(* IEC 61131-3 sources: volt/packages/volt-lsp-iec/test-corpus/bakon-nano/Device/Plc Logic/Application/POUs/LenzeFunctions, 3 files *)

(* ---- SetRef_Axis.pou ---- *)
FUNCTION_BLOCK SetRef_Axis
VAR_INPUT
	I_AxisStatus	: KC_AxisBasicsStatus;
	I_lrHomeTarget	: LREAL;
END_VAR
VAR_OUTPUT
	Q_bRefDone		: BOOL;
	Q_bError		: BOOL;
END_VAR
VAR_IN_OUT
	IQ_CmdSetRef	: BOOL;
	IQ_Axis			: AXIS_REF;
	IQ_uControl_Axis	: KC_AxisBasicsControl;
END_VAR
VAR
	byStepper: BYTE;
	//LenzeECSWriteParameter1: L_DCO_ReadDriveParameter;
	bDone: BOOL;
	bError: BOOL;
	tWait: TON;
	//TestMultiturn: L_SMC_Multiturn;
	SetHomePosition : MC_SetPosition;
END_VAR

%LANGUAGE ST

CASE byStepper OF (*VERVALLEN, KAN NU VIA HOMING IN AXISBASICS: SET HOME -> SM3_Multiturn eronder aanroepen*)

	0:	Q_bRefDone							:=FALSE;
		Q_bError							:=FALSE;

		IF IQ_CmdSetRef
		THEN
			tWait(IN:= FALSE);
			IQ_uControl_Axis.bEnableDrive		:=FALSE;
			bDone								:=FALSE;
			bError								:=FALSE;
			IF NOT I_AxisStatus.bDriveEnabled THEN
				byStepper:=2;
			END_IF
		END_IF

	2:	SetHomePosition.Execute := TRUE;
		IF SetHomePosition.Done OR SetHomePosition.Error THEN
			byStepper := 4;
		END_IF

	4: Q_bRefDone := SetHomePosition.Done;
		Q_bError := SetHomePosition.Error;
		IF NOT IQ_CmdSetRef THEN
			byStepper := 0;
			SetHomePosition.Execute := FALSE;
		END_IF
END_CASE

SetHomePosition(
			Axis	:= IQ_Axis,
			Execute := ,
			Position:= I_lrHomeTarget,
			Relative	:= FALSE,
			Done=> ,
			Busy=> ,
			Error=> ,
			ErrorID=> );

END_FUNCTION_BLOCK

(* ---- XYA_MoveLineair_Bakon.pou ---- *)
(***********************************************************************************
Creation: LENL 		Datum: march 2008		Version: 1.0.0
 ***********************************************************************************
 FUNCTION:

FB for moving XYA in gear mode with a dummy axis. The dummy axis can be positioned or control external

 ***********************************************************************************
Name							Datum				Changes
Kling 							24.03.2009		Implementation

************************************************************************************
NOTE:

***********************************************************************************)

FUNCTION_BLOCK  XYA_MoveLineair_Bakon

VAR
	byStepper: BYTE;
	rMoveX: REAL;
	rMoveY: REAL;
	rMoveA: REAL;
	MC_GearIn_X: MC_GearIn;
	MC_GearIn_Y: MC_GearIn;
	MC_GearIn_A: MC_GearIn;
	MC_GearOut_X: MC_GearOut;
	MC_GearOut_Y: MC_GearOut;
	MC_GearOut_A: MC_GearOut;
	MC_MoveAbsolute_X: MC_MoveAbsolute;
	MC_MoveAbsolute_Y: MC_MoveAbsolute;
	MC_MoveAbsolute_A: MC_MoveAbsolute;
	CalcGearingRatio_X: CalcGearingRatio;
	CalcGearingRatio_Y: CalcGearingRatio;
	CalcGearingRatio_A: CalcGearingRatio;
	CalcGearingRatio_F: CalcGearingRatio;
	CalcGearingRatio_R: CalcGearingRatio;
	MC_MoveAbsolute_Mst: MC_MoveAbsolute;
	MC_SetPosition_Mst: MC_SetPosition;
	CalcMasterSpeedAcc_X: CalcMasterSpeedAcc;
	CalcMasterSpeedAcc_Y: CalcMasterSpeedAcc;
	CalcMasterSpeedAcc_A: CalcMasterSpeedAcc;
	CalcMasterSpeedAcc_F: CalcMasterSpeedAcc;
	CalcMasterSpeedAcc_R: CalcMasterSpeedAcc;
	//MC_Power_Mst: MC_Power;
	rSpeedOverrideOld: REAL;
	MC_Stop_Mst: MC_Stop;
	MC_Halt_X: MC_Halt;
	MC_Halt_Y: MC_Halt;
	MC_Halt_A: MC_Halt;
	rMoveFront: LREAL;
	rMoveRear: LREAL;
END_VAR

VAR_INPUT
	bEnable			: BOOL;
	bPause			: BOOL;
	rMoveMaster		: REAL;
	strTarget			: XYA_Target;
	rSpeedOverride	: REAL:=0.5;
	rAccOverride		: REAL:=0.5;
	bPositionMaster: BOOL;
END_VAR

VAR_IN_OUT
	AxisX		: AXIS_REF;
	AxisY		: AXIS_REF;
	AxisA		: AXIS_REF;
	Master		: AXIS_REF;
END_VAR

VAR_OUTPUT
	bReady		:BOOL;
	bBusy			:BOOL;
	bError			:BOOL;
	nStatus		:INT;
	bAxisAreGearedIn: BOOL;
	bErrorTargetPosInSWLimits: BOOL;
END_VAR

%LANGUAGE ST
	MC_GearIn_X(			Execute:= , 	RatioNumerator:= , 	RatioDenominator:= , 	Acceleration:=AxisX.scPar.MaxAcceleration , 	Deceleration:=AxisX.scPar.MaxAcceleration , 	Master:=Master , 	Slave:=AxisX , 	InGear=> , 	CommandAborted=> , 	Error=> , 	ErrorID=> );
	MC_GearIn_Y(			Execute:=, 		RatioNumerator:= , 	RatioDenominator:= , 	Acceleration:=AxisY.scPar.MaxAcceleration , 	Deceleration:=AxisY.scPar.MaxAcceleration , 	Master:=Master , 	Slave:=AxisY , 	InGear=> , 	CommandAborted=> , 	Error=> , 	ErrorID=> );
	MC_GearIn_A(			Execute:=, 		RatioNumerator:= , 	RatioDenominator:= , 	Acceleration:=AxisA.scPar.MaxAcceleration , 	Deceleration:=AxisA.scPar.MaxAcceleration , 	Master:=Master , 	Slave:=AxisA , 	InGear=> , 	CommandAborted=> , 	Error=> , 	ErrorID=> );
	MC_GearOut_X(			Execute:= , 	Slave:=AxisX , 	Done=> , 	Error=> , 	ErrorID=> );
	MC_GearOut_Y(			Execute:= , 	Slave:=AxisY , 	Done=> , 	Error=> , 	ErrorID=> );
	MC_GearOut_A(			Execute:= , 	Slave:=AxisA , 	Done=> , 	Error=> , 	ErrorID=> );
	MC_MoveAbsolute_X(		Execute:= , 	Position:= , 	Velocity:= , 	Acceleration:= ,	Deceleration:= ,	Direction:= , 	Axis:=AxisX , 	Done=> , 	CommandAborted=> , 	Error=> , 	ErrorID=> );
	MC_MoveAbsolute_Y(		Execute:= , 	Position:= , 	Velocity:= , 	Acceleration:= ,	Deceleration:= ,	Direction:= , 	Axis:=AxisY , 	Done=> , 	CommandAborted=> , 	Error=> , 	ErrorID=> );
	MC_MoveAbsolute_A(		Execute:= , 	Position:= , 	Velocity:= , 	Acceleration:= ,	Deceleration:= ,	Direction:= , 	Axis:=AxisA , 	Done=> , 	CommandAborted=> , 	Error=> , 	ErrorID=> );
	MC_MoveAbsolute_Mst(	Execute:= , 	Position:= , 	Velocity:= , 	Acceleration:= ,	Deceleration:= ,	Direction:=MC_DIRECTION.mcPositiveDirection , 	Axis:=Master , 	Done=> , 	CommandAborted=> , 	Error=> , 	ErrorID=> );
	MC_SetPosition_Mst(		Execute:= ,		Position:=0 , 	Relative:=FALSE , 	Axis:=Master, 	Done=> , 	Error=> , 	ErrorID=> );
	(*MC_Power_Mst(			Enable:=TRUE ,	bRegulatorOn:=TRUE , 	bDriveStart:=TRUE , 	Axis:=Master , 	Status=> ,	Error=> ,	ErrorID=> );*)
	MC_Stop_Mst(			Execute:= ,		Deceleration:=MC_MoveAbsolute_Mst.Deceleration  , 	Axis:=Master , 	Done=> , 	Error=> , 	ErrorID=> );

(*Limiting speed and acc override*)
rSpeedOverride		:=LIMIT(0.01,rSpeedOverride,1);
rAccOverride		:=LIMIT(0.01,rAccOverride,1);

IF NOT bEnable THEN
	byStepper:=0;
	MC_GearIn_X.Execute :=FALSE;
	MC_GearIn_Y.Execute :=FALSE;
	MC_GearIn_A.Execute :=FALSE;
	MC_GearOut_X.Execute:=FALSE;
	MC_GearOut_Y.Execute:=FALSE;
	MC_GearOut_A.Execute:=FALSE;
	MC_MoveAbsolute_X.Execute:=FALSE;
	MC_MoveAbsolute_Y.Execute:=FALSE;
	MC_MoveAbsolute_A.Execute:=FALSE;
	MC_MoveAbsolute_Mst.Execute:=FALSE;
	MC_SetPosition_Mst.Execute:=FALSE;
	MC_Halt_X.Execute:=FALSE;	(* V00.02 *)
	MC_Halt_Y.Execute:=FALSE;	(* V00.02 *)
	MC_Halt_A.Execute:=FALSE;	(* V00.02 *)
	bReady:=FALSE;
	bBusy:=FALSE;
	bError:=FALSE;
	nStatus:=0;
	MC_Stop_Mst.Execute:=FALSE;
	bAxisAreGearedIn		:=FALSE;
	bErrorTargetPosInSWLimits:=FALSE;(*Software-limit error*)
ELSE

CASE byStepper OF
0:		bBusy:=TRUE;

		IF CalcCheckSWLimit_XYA(strTarget, AxisX, AxisY, AxisA) THEN
			byStepper:=200;
		ELSE
			rMoveX:=strTarget.X_Target - AxisX.lrSetPosition ;
			rMoveY:=strTarget.Y_Target - AxisY.lrSetPosition;
			rMoveA:=strTarget.A_Target - AxisA.lrSetPosition;

			rMoveFront := ( strTarget.X_Target + strTarget.Y_Target) - (AxisX.lrSetPosition + AxisY.lrSetPosition );
			rMoveRear := ( strTarget.X_Target - strTarget.Y_Target) - (AxisX.lrSetPosition - AxisY.lrSetPosition );

			IF bPositionMaster THEN
			byStepper:=2;
			ELSE
			byStepper:=10;
			END_IF
		END_IF

2:		MC_SetPosition_Mst.Execute:=TRUE;
		MC_Halt_X.Execute:=TRUE;
		MC_Halt_Y.Execute:=TRUE;
		MC_Halt_A.Execute:=TRUE;

		IF MC_SetPosition_Mst.Done AND MC_Halt_X.Done AND MC_Halt_Y.Done AND MC_Halt_A.Done THEN
		MC_Halt_X.Execute:=FALSE;
		MC_Halt_Y.Execute:=FALSE;
		MC_Halt_A.Execute:=FALSE;
			byStepper:=10;
		END_IF

10:		(*Dummy-axis is the master*)
		CalcGearingRatio_X(	rMoveMaster:=rMoveMaster ,
								rMoveSlave:=rMoveX ,
								nGearNum=> ,
								nGearDenum=>,
								rGearingFactor=> );

		CalcGearingRatio_Y(	rMoveMaster:=rMoveMaster ,
								rMoveSlave:=rMoveY ,
								nGearNum=> ,
								nGearDenum=>,
								rGearingFactor=> );

		CalcGearingRatio_A(	rMoveMaster:=rMoveMaster ,
								rMoveSlave:=rMoveA ,
								nGearNum=> ,
								nGearDenum=>,
								rGearingFactor=> );

		CalcGearingRatio_F(	rMoveMaster:=rMoveMaster ,
								rMoveSlave:=rMoveFront ,
								nGearNum=> ,
								nGearDenum=>,
								rGearingFactor=> );

		CalcGearingRatio_R(	rMoveMaster:=rMoveMaster ,
								rMoveSlave:=rMoveRear ,
								nGearNum=> ,
								nGearDenum=>,
								rGearingFactor=> );

		MC_GearIn_X.RatioNumerator:=CalcGearingRatio_X.nGearNum;
		MC_GearIn_X.RatioDenominator:=INT_TO_UINT( CalcGearingRatio_X.nGearDenum);
		MC_GearIn_X.Execute:=TRUE;

		MC_GearIn_Y.RatioNumerator:=CalcGearingRatio_Y.nGearNum;
		MC_GearIn_Y.RatioDenominator:=INT_TO_UINT( CalcGearingRatio_Y.nGearDenum);
		MC_GearIn_Y.Execute:=TRUE;

		MC_GearIn_A.RatioNumerator:=CalcGearingRatio_A.nGearNum;
		MC_GearIn_A.RatioDenominator:=INT_TO_UINT( CalcGearingRatio_A.nGearDenum);
		MC_GearIn_A.Execute:=TRUE;

		IF MC_GearIn_X.InGear AND MC_GearIn_Y.InGear AND MC_GearIn_A.InGear  THEN
			bAxisAreGearedIn			:=TRUE;
			IF bPositionMaster THEN
			byStepper:=11;
			ELSE
			byStepper:=30;
			END_IF
			rSpeedOverrideOld:=rSpeedOverride;
		END_IF

11:		(*Calculate max-speed and acceleration*)
		CalcMasterSpeedAcc_X(	rGearingRatio:=CalcGearingRatio_X.rGearingFactor  ,	Axis:=AxisX ,	rVelocity=> ,	rAcceleration=> );
		CalcMasterSpeedAcc_Y(	rGearingRatio:=CalcGearingRatio_Y.rGearingFactor  ,	Axis:=AxisY ,	rVelocity=> ,	rAcceleration=> );
		CalcMasterSpeedAcc_A(	rGearingRatio:=CalcGearingRatio_A.rGearingFactor  ,	Axis:=AxisA ,	rVelocity=> ,	rAcceleration=> );
		CalcMasterSpeedAcc_F(	rGearingRatio:=CalcGearingRatio_F.rGearingFactor , Axis := Front_Axis, rVelocity=>, rAcceleration=>);
		CalcMasterSpeedAcc_R(	rGearingRatio:=CalcGearingRatio_R.rGearingFactor , Axis := Rear_Axis, rVelocity=>, rAcceleration=>);
		(*Move X to target*)
		MC_MoveAbsolute_Mst.Position:=rMoveMaster;
		MC_MoveAbsolute_Mst.Velocity:=MIN(CalcMasterSpeedAcc_F.rVelocity,MIN(CalcMasterSpeedAcc_R.rVelocity, MIN(MIN(CalcMasterSpeedAcc_X.rVelocity, CalcMasterSpeedAcc_Y.rVelocity), CalcMasterSpeedAcc_A.rVelocity))) * rSpeedOverride;
		MC_MoveAbsolute_Mst.Acceleration:=MIN(CalcMasterSpeedAcc_F.rAcceleration,MIN(CalcMasterSpeedAcc_R.rAcceleration,MIN(MIN(CalcMasterSpeedAcc_X.rAcceleration, CalcMasterSpeedAcc_Y.rAcceleration), CalcMasterSpeedAcc_A.rAcceleration))) * rAccOverride ;
		MC_MoveAbsolute_Mst.Deceleration:=MC_MoveAbsolute_Mst.Acceleration;
		MC_MoveAbsolute_Mst.Execute:=TRUE;

		IF MC_MoveAbsolute_Mst.Done THEN
			MC_MoveAbsolute_Mst.Execute:=FALSE;
			byStepper:=80;
		END_IF

		(*Restart positioning if SpeedOverride  changes*)
		IF rSpeedOverride <> rSpeedOverrideOld THEN
					MC_MoveAbsolute_Mst.Execute:=FALSE;
					rSpeedOverrideOld:=rSpeedOverride;
					byStepper:=13;
		END_IF

		(*Pause*)
		IF bPause THEN
			byStepper:=20;
			MC_Stop_Mst.Execute:=TRUE;
			MC_MoveAbsolute_Mst.Execute:=FALSE;
		END_IF

13:		(*Restart*)
		byStepper:=11;

20:		(*Restart after pause*)
		IF NOT bPause THEN
			MC_Stop_Mst.Execute:=FALSE;
			byStepper:=11;
		END_IF

30:		IF Master.lrActPosition >= (rMoveMaster - 0.1) THEN	(*This is important! Axes are currently geared in, so will follow the movement of the Master axis! gear at when the master made a complete move!*)
			byStepper:=80;
		END_IF

80:		(*Gear-out*)
		MC_GearOut_X.Execute:=TRUE;
		MC_GearOut_Y.Execute:=TRUE;
		MC_GearOut_A.Execute:=TRUE;

		IF MC_GearOut_X.Done AND  MC_GearOut_Y.Done AND  MC_GearOut_A.Done THEN
			MC_GearOut_X.Execute:=FALSE;
			MC_GearOut_Y.Execute:=FALSE;
			MC_GearOut_A.Execute:=FALSE;
			MC_GearIn_X.Execute:=FALSE;
			MC_GearIn_Y.Execute:=FALSE;
			MC_GearIn_A.Execute:=FALSE;
			bAxisAreGearedIn		:=FALSE;
			byStepper:=90;
		END_IF

90:		(*single axis-movement*)
			MC_MoveAbsolute_X.Position:=strTarget.X_Target;
			MC_MoveAbsolute_X.Velocity:=AxisX.scPar.MaxVelocity;
			MC_MoveAbsolute_X.Acceleration:=AxisX.scPar.MaxAcceleration;
			MC_MoveAbsolute_X.Deceleration:=AxisX.scPar.MaxAcceleration;	//Was fSWMaxDeceleration in old motion
			MC_MoveAbsolute_X.Direction:=MC_DIRECTION.mcShortestWay;
			MC_MoveAbsolute_X.Execute:=TRUE;

			MC_MoveAbsolute_Y.Position:=strTarget.Y_Target;
			MC_MoveAbsolute_Y.Velocity:=AxisY.scPar.MaxVelocity;
			MC_MoveAbsolute_Y.Acceleration:=AxisY.scPar.MaxAcceleration;
			MC_MoveAbsolute_Y.Deceleration:=AxisY.scPar.MaxAcceleration;	//Was fSWMaxDeceleration in old motion
			MC_MoveAbsolute_Y.Direction:=MC_DIRECTION.mcShortestWay;
			MC_MoveAbsolute_Y.Execute:=TRUE;

			MC_MoveAbsolute_A.Position:=strTarget.A_Target;
			MC_MoveAbsolute_A.Velocity:=AxisA.scPar.MaxVelocity;
			MC_MoveAbsolute_A.Acceleration:=AxisA.scPar.MaxAcceleration;
			MC_MoveAbsolute_A.Deceleration:=AxisA.scPar.MaxAcceleration;	//Was fSWMaxDeceleration in old motion
			MC_MoveAbsolute_A.Direction:=MC_DIRECTION.mcShortestWay;
			MC_MoveAbsolute_A.Execute:=TRUE;

			IF MC_MoveAbsolute_X.Done AND MC_MoveAbsolute_Y.Done AND MC_MoveAbsolute_A.Done THEN
				byStepper:=100;
			END_IF

100:		(*Ready*)
			bBusy:=FALSE;
			bReady:=TRUE;

200:		bErrorTargetPosInSWLimits:=TRUE;(*Software-limit error*)
			;
END_CASE

MC_Halt_X(
	Execute:= ,
	Deceleration:= 100,
	Axis:=AxisX ,
	Done=> ,
	CommandAborted=> ,
	Error=> ,
	ErrorID=> );

MC_Halt_Y(
	Execute:= ,
	Deceleration:= 100,
	Axis:=AxisY ,
	Done=> ,
	CommandAborted=> ,
	Error=> ,
	ErrorID=> );

MC_Halt_A(
	Execute:= ,
	Deceleration:= 100,
	Axis:=AxisA ,
	Done=> ,
	CommandAborted=> ,
	Error=> ,
	ErrorID=> );
END_IF

bError:=		MC_GearIn_X.Error OR MC_GearIn_Y.Error OR MC_GearIn_A.Error OR MC_GearOut_X.Error OR MC_GearOut_Y.Error OR MC_GearOut_A.Error OR
				MC_MoveAbsolute_X.Error OR MC_MoveAbsolute_Y.Error OR MC_MoveAbsolute_A.Error OR MC_MoveAbsolute_Mst.Error OR MC_SetPosition_Mst.Error (*OR MC_Power_Mst.Error TODO: AxisBasics Status*) OR (byStepper =200);

END_FUNCTION_BLOCK

(* ---- ModusRondVierkant.pou ---- *)
(***********************************************************************************
Creation: LENL 		Datum: juli 2012		Version: 1.0.0
 ***********************************************************************************
 FUNCTION:

Cutting round or square products with XYAZ axis

 ***********************************************************************************
Name							Datum				Changes
Kling 							20.07.2012			Implementation		Version 1.0.0

************************************************************************************
NOTE:

***********************************************************************************)
PROGRAM ModusRondVierkant

VAR
	MC_SetPosition1					: MC_SetPosition;
	XYA_MoveLineair_Bakon1			: XYA_MoveLineair_Bakon;
	byStepper						: BYTE;
	nLineNumber						: INT;
	nCount							: INT;
	R_TRIG1							: R_TRIG;
	byStepperOLd1					: BYTE;
	rZactPos						: REAL;
	rParaAccTime					: REAL:=0.1;
	Check_Table1					: Check_Table_V2;
	MC_MoveAbsoluteZ				: MC_MoveAbsolute;
	fRampJerkDummyAxis				: LREAL;
	rSlowPart						: REAL;
	nCleanCountProd					: INT;
	nCleanCountCuts					: INT;
	bLastCut						: BOOL;
	MC_HaltZ						: MC_Halt;
	rVelocityZ						: LREAL;
	rAccelerationZ					: LREAL;
	bCrashDetectWasOK				: BOOL;
END_VAR

VAR_INPUT
	I_bEnable						: BOOL;
	I_bStartXYA						: BOOL;
	I_bStartZ						: BOOL;
	I_TableCheckSensor				: BOOL;
	I_bTestMode						: BOOL;
	//I_bCleanRequest				: BOOL;
	I_strParameters					: strRondVierkantParameters;
	I_rSpeedOverride				: REAL:=0.5;
	I_rAccOverride					: REAL:=0.5;
	I_rX_InfeedPosition				: REAL;
	I_rY_InfeedPrePosition			: REAL;
	I_rY_InfeedPosition				: REAL;
	I_rA_EndTarget					: REAL;
END_VAR

VAR_IN_OUT
	IQ_AxisX						:AXIS_REF;
	IQ_AxisY						:AXIS_REF;
	IQ_AxisA						:AXIS_REF;
	IQ_AxisZ						:AXIS_REF;
	IQ_AxisDummy					:AXIS_REF;
	IQ_strTarget					: ARRAY [1..C_wNumberOfMotionObjects] OF XYA_Target;
END_VAR

VAR_OUTPUT
	Q_bReady						: BOOL;
	Q_bLastCutReadyZOutOfProduct	: BOOL;
	Q_bErrorTargetPosInSWLimits		: BOOL;
	Q_bErrorAccDeccZ				: BOOL;
	Q_bErrorSpeedZToHigh			: BOOL;
	Q_nActLineNumber				: INT;
	Q_byCounter						: BYTE;
END_VAR

%LANGUAGE ST
MC_MoveAbsoluteZ(
	Execute:= ,
	Position:= ,
	Velocity:= ,
	Acceleration:= ,
	Deceleration:= ,
	Direction:=MC_DIRECTION.mcShortestWay ,
	Axis:=IQ_AxisZ ,
	Done=> ,
	CommandAborted=> ,
	Error=> ,
	ErrorID=> );

MC_HaltZ(
	Execute 	:= ,
	Deceleration:= IQ_AxisZ.scPar.MaxAcceleration,	//Was fSWMaxDeceleration in old motion
	Jerk		:= ,
	Axis		:= IQ_AxisZ,
	Done 	=> ,
	Busy 	=> ,
	CommandAborted =>,
	Error	=> ,
	ErrorID => );

MC_SetPosition1(
	Execute:= ,
	Position:=0 ,
	Relative:=FALSE ,
	Axis:=IQ_AxisDummy ,
	Done=> ,
	Error=> ,
	ErrorID=> );

XYA_MoveLineair_Bakon1(
	bEnable:= ,
	bPause:= ,
	rMoveMaster		:=359 ,
	strTarget:= ,
	rSpeedOverride	:=I_rSpeedOverride * rSlowPart,
	rAccOverride		:=I_rAccOverride ,
	bPositionMaster	:= ,
	AxisX				:=IQ_AxisX ,
	AxisY				:=IQ_AxisY ,
	AxisA				:=IQ_AxisA ,
	Master				:=IQ_AxisDummy ,
	bReady=> ,
	bBusy=> ,
	bErrorTargetPosInSWLimits=>Q_bErrorTargetPosInSWLimits ,
	nStatus=> );

Check_Table1(
	I_bStartCheck			:= ,				(* Start check when table moves from infeed position to first cutting position *)
	I_bSensor				:= I_TableCheckSensor,
	I_bTestModus			:= I_bTestMode,
	I_nProdTypeSelection	:= SEL(g_HMI_MachCommand.bScanMode, g_HMI_RCP_Parameters.nProductType,-1),
	I_nPartsRoundLeft		:= g_HMI_RCP_Parameters.nPartsRound,
	I_nPartsRoundRight		:= g_HMI_RCP_Parameters.nPartsRoundRight,
	I_rActualPositionY		:= g_uStatus_Y_Axis.lrActPosition,
	Q_TabelCheckOK			=> );

Q_nActLineNumber						:=nLineNumber;

(*Crash detectie sensor*)
IF 	NOT g_uStatus_Z_Axis.bDigIn1
	AND g_uStatus_Z_Axis.lrActPosition < I_strParameters.strZasParameters.rCrashCheckHeight
	AND (byStepper = 9 OR byStepper = 10)
	//AND g_HMI_RCP_Parameters.bCutWasteFirst
	AND gMachConfig.bCrashDetection
	THEN
		g_sMACH.ERR.bCrashDetected := TRUE;
END_IF

IF NOT I_bEnable THEN
	MC_MoveAbsoluteZ.Execute		:=FALSE;
	MC_Setposition1.Execute			:=FALSE;
	XYA_MoveLineair_Bakon1.bEnable	:=FALSE;
	byStepper						:=0;
	nLineNumber						:=C_wNumberOfMotionObjects + 100;
	nCount							:=0;
	Q_byCounter						:=0;
	R_TRIG1(CLK:=FALSE);
	Q_bReady						:=FALSE;
	Q_bLastCutReadyZOutOfProduct	:=FALSE;
	Q_bErrorSpeedZToHigh			:=FALSE;
	Q_bErrorAccDeccZ				:=FALSE;
	g_bUS_EnableRV					:=FALSE;
	Check_Table1.I_bStartCheck		:=FALSE;
	rSlowPart						:= 1;
	MC_HaltZ.Execute				:= FALSE;
	bCrashDetectWasOK := FALSE;
ELSE

	(*actuele jerk time bij onderbreking van beweging*)
	fRampJerkDummyAxis					:=IQ_AxisDummy.scPar.JerkErrorStop;

(*	R_TRIG1(CLK:=(IQ_AxisZ.lrActPosition <= (I_strParameters.strZasParameters.rBottomZPos - I_strParameters.strZasParameters.rProductHeigt)) AND
				(IQ_AxisZ.lrActPosition >= (I_strParameters.strZasParameters.rBottomZPos - I_strParameters.strZasParameters.rProductHeigt - 10))); *)
	R_TRIG1(CLK:=(IQ_AxisZ.lrActPosition <= (I_strParameters.strZasParameters.rAboveProductPos)) AND
				(IQ_AxisZ.lrActPosition >= (I_strParameters.strZasParameters.rAboveProductPos - 10)));

	IF R_TRIG1.Q THEN
		byStepperOld1					:=byStepper;
		rZactPos							:=IQ_AxisZ.lrActPosition;
	END_IF

	CASE byStepper OF
	0:	IF I_bStartXYA THEN
			Q_bLastCutReadyZOutOfProduct	:=FALSE;
			Q_bReady							:=FALSE;
			nLineNumber						:=C_wNumberOfMotionObjects + 100;
			byStepper							:=2;
		END_IF

	(*check position table for XYA*)
	2:	FOR nCount:=C_wNumberOfMotionObjects TO 1 BY -1 DO
			IF (IQ_strTarget[nCount].X_Target >= 0) AND (IQ_strTarget[nCount].Y_Target >= 0) AND (IQ_strTarget[nCount].A_Target >= 0) THEN
				nLineNumber:=nCount;
			END_IF
		END_FOR
		IF nLineNumber = (C_wNumberOfMotionObjects + 100) THEN
			Q_bReady := TRUE;
			byStepper:=0;
		ELSE
			byStepper:=3;
		END_IF

	(* Go to the left in order to start the table check*)
	3:	XYA_MoveLineair_Bakon1.strTarget.X_Target:=C_rTargetX_TableCheck;
		XYA_MoveLineair_Bakon1.strTarget.Y_Target:=40;		(* @TODO: Mach Par ? *)
		XYA_MoveLineair_Bakon1.strTarget.A_Target:=IQ_strTarget[nLineNumber].A_Target;

		XYA_MoveLineair_Bakon1.bPositionMaster	:=TRUE;
		XYA_MoveLineair_Bakon1.bEnable			:=TRUE;

		IF XYA_MoveLineair_Bakon1.bReady THEN
			XYA_MoveLineair_Bakon1.bPositionMaster:=FALSE;
			XYA_MoveLineair_Bakon1.bEnable	:=FALSE;
			rSlowPart				:= 0.7;
			bCrashDetectWasOK := FALSE;
			byStepper				:=4;
		END_IF

	(* Go to the rear and start the table check*)
	4:	XYA_MoveLineair_Bakon1.strTarget.X_Target:=C_rTargetX_TableCheck;
		XYA_MoveLineair_Bakon1.strTarget.Y_Target:=SEL(gMachConfig.bXL, 265,390);		(* @TODO: Mach Par ? *)
		XYA_MoveLineair_Bakon1.strTarget.A_Target:=IQ_strTarget[nLineNumber].A_Target;

		XYA_MoveLineair_Bakon1.bPositionMaster	:=TRUE;
		XYA_MoveLineair_Bakon1.bEnable			:=TRUE;

		Check_Table1.I_bStartCheck			:= TRUE;		(* Check if table correspondents with recipe *)
		IF Check_Table1.Q_bCrashDetectionOK THEN
			bCrashDetectWasOK := TRUE;
		END_IF
		IF XYA_MoveLineair_Bakon1.bReady THEN
			IF	Check_Table1.Q_TabelCheckOK AND bCrashDetectWasOK THEN
				Check_Table1.I_bStartCheck				:= FALSE;
				XYA_MoveLineair_Bakon1.bPositionMaster	:=FALSE;
				XYA_MoveLineair_Bakon1.bEnable			:=FALSE;
				rSlowPart					:= 1.0;
				bCrashDetectWasOK := FALSE;
				byStepper					:=5;
			ELSE
				g_sMACH.ERR.bCrashDetectFault 	:= NOT bCrashDetectWasOK;
				g_sMACH.ERR.bWrongTable			:= NOT Check_Table1.Q_TabelCheckOK;
				Check_Table1.I_bStartCheck		:= FALSE;
			END_IF
		END_IF

	(*start first positioning of XYA*)
	5:	XYA_MoveLineair_Bakon1.strTarget:=IQ_strTarget[nLineNumber];
		XYA_MoveLineair_Bakon1.bPositionMaster	:=TRUE;
		XYA_MoveLineair_Bakon1.bEnable			:=TRUE;

		IF XYA_MoveLineair_Bakon1.bReady THEN
			XYA_MoveLineair_Bakon1.bPositionMaster:=FALSE;
			XYA_MoveLineair_Bakon1.bEnable	:=FALSE;
			(*nLineNumber					:=nLineNumber+1; *)
			byStepper						:=6;
		END_IF

	(*wait for startsignal Z*)
	6:	IF I_bStartZ THEN
			byStepper						:=8;
		END_IF

	(*set dummy to zero pos*)
	8:	MC_Setposition1.Execute			:=TRUE;
		IF MC_Setposition1.Done THEN
			MC_Setposition1.Execute	:=FALSE;
			IF IQ_strTarget[nLineNumber].bCrashDetectCheck AND g_uStatus_Z_Axis.lrActPosition < I_strParameters.strZasParameters.rAboveProductPos-8 THEN //AC Aanpassing 24-07-2018
				byStepper						:=9;
			ELSE
				byStepper						:=10;
			END_IF
		END_IF

	(*In between step for quick start i.c.w. edge detection*)
	9:	MC_MoveAbsoluteZ.Position		:= I_strParameters.strZasParameters.rCrashCheckHeight - 10;
		rVelocityZ	:= I_strParameters.strZasParameters.rCuttingSpeedDown;
		rAccelerationZ	:= I_strParameters.strZasParameters.rCuttingSpeedDown / rParaAccTime;
		MC_MoveAbsoluteZ.Velocity		:=rVelocityZ;
		MC_MoveAbsoluteZ.Acceleration	:=rAccelerationZ;
		MC_MoveAbsoluteZ.Deceleration	:=MC_MoveAbsoluteZ.Acceleration;
		MC_MoveAbsoluteZ.Execute		:= NOT g_sMACH.ERR.bCrashDetected; // TRUE;
		IF MC_MoveAbsoluteZ.Done OR g_sMACH.ERR.bCrashDetected THEN		(* Crash detection *)
			MC_MoveAbsoluteZ.Execute		:=FALSE;
			IF g_sMACH.ERR.bCrashDetected THEN	(* Crash detection *)
				MC_HaltZ.Execute	:= TRUE;
				IF MC_HaltZ.Done THEN
					MC_HaltZ.Execute	:= FALSE;
					byStepper	:= 12;
				END_IF
			ELSE
				byStepper		:= 10;
			END_IF
		END_IF
	(*z-as to bottom pos*)
	10:
		MC_MoveAbsoluteZ.Position		:=SEL(IQ_strTarget[nLineNumber].bCrashDetectCheck, I_strParameters.strZasParameters.rBottomZPos, I_strParameters.strZasParameters.rCrashCheckHeight);
		IF g_HMI_MachCommand.bScanMode THEN
			rVelocityZ		:= 480;
			rAccelerationZ	:= 480 / rParaAccTime;
		ELSIF IQ_strTarget[nLineNumber].bCrashDetectCheck THEN  // Langzamere snelheid tijdens crash check
			rVelocityZ	:= g_HMI_MCH_Parameters.rSpeedZ_CrashDetect;
			rAccelerationZ	:= 50 / rParaAccTime;
		ELSE
			rVelocityZ	:= I_strParameters.strZasParameters.rCuttingSpeedDown;
			rAccelerationZ	:= I_strParameters.strZasParameters.rCuttingSpeedDown / rParaAccTime;
		END_IF
		MC_MoveAbsoluteZ.Velocity		:=rVelocityZ;
		MC_MoveAbsoluteZ.Acceleration	:=rAccelerationZ;
		MC_MoveAbsoluteZ.Deceleration	:=MC_MoveAbsoluteZ.Acceleration;
		MC_MoveAbsoluteZ.Execute		:= NOT g_sMACH.ERR.bCrashDetected; // TRUE;
		IF MC_MoveAbsoluteZ.Done OR g_sMACH.ERR.bCrashDetected THEN		(* Crash detection *)
			MC_MoveAbsoluteZ.Execute		:=FALSE;
			IF g_sMACH.ERR.bCrashDetected THEN	(* Crash detection *)
				MC_HaltZ.Execute	:= TRUE;
				IF MC_HaltZ.Done THEN
					MC_HaltZ.Execute	:= FALSE;
					byStepper	:= 12;
				END_IF
			ELSE
				byStepper		:= 12;
			END_IF
		END_IF

	(*z-as to above or top product pos*)
	12:
		IF		((IQ_strTarget[nLineNumber+1].X_Target = -50)	(* controleer de volgende positie *)
			AND	(IQ_strTarget[nLineNumber+1].Y_Target = -50)
			AND	(IQ_strTarget[nLineNumber+1].A_Target = -50))
			OR	g_sMACH.ERR.bCrashDetected
		THEN
			MC_MoveAbsoluteZ.Position		:=I_strParameters.strZasParameters.rTopZPos;
			MC_MoveAbsoluteZ.Velocity		:=SEL(g_HMI_MachCommand.bScanMode,	I_strParameters.strZasParameters.rCuttingSpeedUp,480);//I_strParameters.strZasParameters.rCuttingSpeedUp;			(* Std V02.09, was voorheen rSpeedOutProduct *)
			IF R_TRIG1.Q THEN
				Q_bLastCutReadyZOutOfProduct		:=TRUE;
			END_IF
		ELSE
			MC_MoveAbsoluteZ.Position		:=I_strParameters.strZasParameters.rAboveProductPos;
			MC_MoveAbsoluteZ.Velocity		:=SEL(g_HMI_MachCommand.bScanMode,	I_strParameters.strZasParameters.rCuttingSpeedUp,480);//I_strParameters.strZasParameters.rCuttingSpeedUp;
		END_IF

		MC_MoveAbsoluteZ.Acceleration	:=(MC_MoveAbsoluteZ.Velocity / rParaAccTime);
		MC_MoveAbsoluteZ.Deceleration	:=MC_MoveAbsoluteZ.Acceleration;
		MC_MoveAbsoluteZ.Execute		:=TRUE;
		IF		MC_MoveAbsoluteZ.Done
			//OR	R_TRIG1.Q
		THEN
				Q_byCounter					:=Q_byCounter + BOOL_TO_BYTE(NOT g_sMACH.ERR.bCrashDetected);
				IQ_strTarget[nLineNumber].X_Target	:=-50;
				IQ_strTarget[nLineNumber].Y_Target	:=-50;
				IQ_strTarget[nLineNumber].A_Target	:=-50;
				nLineNumber					:=nLineNumber+1;
				bLastCut	:= 	(IQ_strTarget[nLineNumber].X_Target = -50)	// Laatste snede
							AND	(IQ_strTarget[nLineNumber].Y_Target = -50)
							AND	(IQ_strTarget[nLineNumber].A_Target = -50);
				IF	bLastCut THEN
					nCleanCountProd	:= nCleanCountProd + 1;	// ophogen productteller
				END_IF
				nCleanCountCuts	:= nCleanCountCuts + 1; // ophogen snijteller
				IF g_HMI_RCP_Parameters.nCleanAfterNProd = 0 THEN
					nCleanCountCuts := 0;
					nCleanCountProd := 0;
				END_IF
				byStepper					:=14;
		END_IF

	(*start next positioning of XYA or Cleaning cycle or Last cut *)
	14:	(* Clean request *)
		IF		((g_HMI_MachCommand.CMD.bCleanKnifeRequest AND (g_HMI_RCP_Parameters.nCleanProdOrCuts = nCleanAfterProducts) AND bLastCut)
			OR	(g_HMI_MachCommand.CMD.bCleanKnifeRequest AND (g_HMI_RCP_Parameters.nCleanProdOrCuts = nCleanAfterCuts))
			OR  ((nCleanCountProd >= g_HMI_RCP_Parameters.nCleanAfterNProd) AND (g_HMI_RCP_Parameters.nCleanAfterNProd <> 0) AND (g_HMI_RCP_Parameters.nCleanProdOrCuts = nCleanAfterProducts))
			OR  ((nCleanCountCuts >= g_HMI_RCP_Parameters.nCleanAfterNProd) AND (g_HMI_RCP_Parameters.nCleanAfterNProd <> 0) AND (g_HMI_RCP_Parameters.nCleanProdOrCuts = nCleanAfterCuts)))
			AND	gMachConfig.bCleaningUnit
			AND NOT g_sMACH.ERR.bCrashDetected
		THEN
			nCleanCountProd	:= 0;
			nCleanCountCuts	:= 0;
			g_bCleanRequest	:= TRUE;
		END_IF

		(*start next positioning of XYA or Cleaning cycle or Last cut *)
		IF		bLastCut
			OR	g_bCleanRequest
			OR	g_sMACH.ERR.bCrashDetected
		THEN
			MC_MoveAbsoluteZ.Velocity	:=SEL(g_HMI_MachCommand.bScanMode,	I_strParameters.strZasParameters.rCuttingSpeedUp,480);//I_strParameters.strZasParameters.rCuttingSpeedUp;I_strParameters.strZasParameters.rSpeedOutProduct;			(* Std V02.09, snelheid boven product hoger *)
			MC_MoveAbsoluteZ.Execute	:=FALSE;						(* Std V02.09, snelheid boven product hoger *)
			IF	(bLastCut AND NOT g_bCleanRequest) OR g_sMACH.ERR.bCrashDetected THEN
				byStepper					:=20;
			ELSE
				g_bCleanRequest	:= FALSE;
				g_HMI_MachCommand.CMD.bCleanKnifeRequest	:= FALSE;
				g_bSUB_CleanKnifeStart		:= TRUE;
				byStepper					:=16;
			END_IF
		ELSE
			MC_MoveAbsoluteZ.Execute	:=FALSE;
			XYA_MoveLineair_Bakon1.strTarget	:= IQ_strTarget[nLineNumber];
			XYA_MoveLineair_Bakon1.bPositionMaster	:=TRUE;
			XYA_MoveLineair_Bakon1.bEnable			:=TRUE;
			IF XYA_MoveLineair_Bakon1.bReady THEN
				XYA_MoveLineair_Bakon1.bPositionMaster:=FALSE;
				XYA_MoveLineair_Bakon1.bEnable	:=FALSE;
				(*IQ_strTarget[nLineNumber].X_Target	:=-50;
				IQ_strTarget[nLineNumber].Y_Target	:=-50;
				IQ_strTarget[nLineNumber].A_Target	:=-50;
				nLineNumber							:=nLineNumber+1; *)
				byStepper						:=8;
			END_IF
		END_IF

	(* Wait for Cleaning cycle done *)
	16:
	IF	g_bSUB_CleanKnifeDone
	THEN
		g_bSUB_CleanKnifeStart			:= FALSE;
	END_IF

	IF NOT g_bSUB_CleanKnifeStart THEN
		IF	bLastCut THEN
			byStepper					:=20;
		ELSE
			XYA_MoveLineair_Bakon1.strTarget	:= IQ_strTarget[nLineNumber];
			XYA_MoveLineair_Bakon1.bPositionMaster	:=TRUE;
			XYA_MoveLineair_Bakon1.bEnable			:=TRUE;
			IF XYA_MoveLineair_Bakon1.bReady THEN
				XYA_MoveLineair_Bakon1.bPositionMaster:=FALSE;
				XYA_MoveLineair_Bakon1.bEnable	:=FALSE;
				byStepper						:=8;
			END_IF
		END_IF
	END_IF

	(*pos back XYA to operator place pre position *)
	20:
		MC_MoveAbsoluteZ.Execute	:= TRUE;						(* Std V02.09, snelheid boven product hoger *)
		XYA_MoveLineair_Bakon1.strTarget.X_Target:=I_rX_InfeedPosition;
		XYA_MoveLineair_Bakon1.strTarget.Y_Target:=I_rY_InfeedPrePosition;
		XYA_MoveLineair_Bakon1.strTarget.A_Target:=0;	// Ivm beperkte hoogte Nano mes altijd naar 0 graden!!   I_rA_EndTarget;
		XYA_MoveLineair_Bakon1.bPositionMaster	:=TRUE;
		XYA_MoveLineair_Bakon1.bEnable			:=TRUE;
		IF XYA_MoveLineair_Bakon1.bReady THEN
			XYA_MoveLineair_Bakon1.bPositionMaster	:=FALSE;
			XYA_MoveLineair_Bakon1.bEnable			:=FALSE;
			//nCleanCount					:= nCleanCount + 1;
			byStepper								:=22;
		END_IF

	(*pos back XYA to operator place position *)
	22:
		rSlowPart			:= 0.25;
		XYA_MoveLineair_Bakon1.strTarget.X_Target:=I_rX_InfeedPosition;

		IF I_bTestMode THEN
			XYA_MoveLineair_Bakon1.strTarget.Y_Target:=I_rY_InfeedPrePosition;
		ELSE
			XYA_MoveLineair_Bakon1.strTarget.Y_Target:=I_rY_InfeedPosition;
		END_IF
		IF	MC_MoveAbsoluteZ.Done THEN
			MC_MoveAbsoluteZ.Execute	:=FALSE;
			XYA_MoveLineair_Bakon1.strTarget.A_Target:=I_rA_EndTarget;
			XYA_MoveLineair_Bakon1.bPositionMaster	:=TRUE;
			XYA_MoveLineair_Bakon1.bEnable			:=TRUE;
		END_IF
		IF XYA_MoveLineair_Bakon1.bReady
		THEN
			XYA_MoveLineair_Bakon1.bPositionMaster	:=FALSE;
			XYA_MoveLineair_Bakon1.bEnable			:=FALSE;
			rSlowPart								:=1;
			Q_bReady								:=TRUE;
			Q_byCounter								:=0;
			byStepper								:=0;
		END_IF

	END_CASE

	IF (MC_MoveAbsoluteZ.Acceleration > IQ_AxisZ.scPar.MaxAcceleration) OR
		(MC_MoveAbsoluteZ.Acceleration > IQ_AxisZ.scPar.MaxAcceleration) THEN
		Q_bErrorAccDeccZ:=TRUE;
	ELSE
		Q_bErrorAccDeccZ:=FALSE;
	END_IF
	IF (I_strParameters.strZasParameters.rSpeedOutProduct > IQ_AxisZ.scPar.MaxVelocity) OR
		(I_strParameters.strZasParameters.rCuttingSpeedDown > IQ_AxisZ.scPar.MaxVelocity) OR
		(I_strParameters.strZasParameters.rCuttingSpeedUp > IQ_AxisZ.scPar.MaxVelocity) THEN
		Q_bErrorSpeedZToHigh:=TRUE;
	ELSE
		Q_bErrorSpeedZToHigh:=FALSE;
	END_IF

	g_bUS_EnableRV	:= 		((IQ_AxisZ.lrActPosition >= (I_strParameters.strZasParameters.rBottomZPos - g_HMI_RCP_Parameters.rUSHeightStart)) AND byStepper = 10)
						OR	((IQ_AxisZ.lrActPosition >= (I_strParameters.strZasParameters.rBottomZPos - g_HMI_RCP_Parameters.rUSHeightStop)) AND byStepper = 12);

END_IF

END_PROGRAM
